Staubli VAL3: Atan2.pgx

public program Atan2(num y, num x, num& angle)
begin
  //双变量反正切函数atan2(x,y)
  if x>0
    angle=atan(y/x)
  elseIf y>=0 and x<0
    angle=atan(y/x)+180
  elseIf y<0 and x<0
    angle=atan(y/x)-180
  elseIf y>0 and x==0
    angle=90
  elseIf y<0 and x==0
    angle=-90
  elseIf y==0 and x==0
    //Undefined
  endIf
end
